(* IEC 61131-3 sources: ironplc/compiler/ironplc-cli/resources/test/set, 1 file *)

(* ---- first_steps_configuration.st ---- *)
CONFIGURATION config
  VAR_GLOBAL CONSTANT
    ResetCounterValue : INT := 17;
  END_VAR

  RESOURCE resource1 ON PLC
    TASK plc_task(INTERVAL := T#100ms,PRIORITY := 1);
    PROGRAM plc_task_instance WITH plc_task : plc_prg;
  END_RESOURCE
END_CONFIGURATION
